(* IEC 61131-3 sources: kns-pump-station/tests/POUs/Station/FB_Protections_Test, 24 files *)

(* ---- DryRunAndEmergencyBothDryRunWins.method.decl.st ---- *)
// 04 §10.2: сухой ход и аварийный уровень одновременно — оба признака (старшинство сухого хода —
// FB_ControlSelector), по поплавкам LS103 останавливает откачку
METHOD PRIVATE DryRunAndEmergencyBothDryRunWins
VAR
    fbDut  : FB_Protections;            // ФБ под тестом
    fbTime : PL.FB_FakeTime;            // подменное время, старт 1 ч
    stCfg  : ST_StationCfg;             // уставки по умолчанию (tLdev 30 с, tLtRecover 30 с, tDryRelease 60 с)
    fbSink : FB_FakeEventSink;          // подменный журнал
END_VAR

(* ---- DryRunByFloat.method.decl.st ---- *)
// 04 §10.1, PMI-19: поплавок LS103 сработал — сухой ход сразу (защита срабатывает до проверки согласования)
METHOD PRIVATE DryRunByFloat
VAR
    fbDut  : FB_Protections;            // ФБ под тестом
    fbTime : PL.FB_FakeTime;            // подменное время, старт 1 ч
    stCfg  : ST_StationCfg;             // уставки по умолчанию (tLdev 30 с, tLtRecover 30 с, tDryRelease 60 с)
    fbSink : FB_FakeEventSink;          // подменный журнал
END_VAR

(* ---- DryRunByLtLl.method.decl.st ---- *)
// 04 §10.1, PMI-18: LL по годному уровнемеру — сухой ход
METHOD PRIVATE DryRunByLtLl
VAR
    fbDut  : FB_Protections;            // ФБ под тестом
    fbTime : PL.FB_FakeTime;            // подменное время, старт 1 ч
    stCfg  : ST_StationCfg;             // уставки по умолчанию (tLdev 30 с, tLtRecover 30 с, tDryRelease 60 с)
    fbSink : FB_FakeEventSink;          // подменный журнал
END_VAR

(* ---- DryRunReleaseAboveL.method.decl.st ---- *)
// 04 §10.1, PMI-18: снятие сухого хода — LS103 не сработал, нет LL и уровень выше L (по флагу L уровнемера)
METHOD PRIVATE DryRunReleaseAboveL
VAR
    fbDut  : FB_Protections;            // ФБ под тестом
    fbTime : PL.FB_FakeTime;            // подменное время, старт 1 ч
    stCfg  : ST_StationCfg;             // уставки по умолчанию (tLdev 30 с, tLtRecover 30 с, tDryRelease 60 с)
    fbSink : FB_FakeEventSink;          // подменный журнал
END_VAR

(* ---- DryRunReleaseWithoutLtAfterTDryRelease.method.decl.st ---- *)
// 04 §10.1, §11, PMI-19: без уровнемера сухой ход снимается, когда LS103 снят дольше tDryRelease = 60 с (не
// раньше)
METHOD PRIVATE DryRunReleaseWithoutLtAfterTDryRelease
VAR
    fbDut  : FB_Protections;            // ФБ под тестом
    fbTime : PL.FB_FakeTime;            // подменное время, старт 1 ч
    stCfg  : ST_StationCfg;             // уставки по умолчанию (tLdev 30 с, tLtRecover 30 с, tDryRelease 60 с)
    fbSink : FB_FakeEventSink;          // подменный журнал
END_VAR

(* ---- EmergencyByFloatAndByHh.method.decl.st ---- *)
// 04 §10.2, PMI-20, PMI-23: аварийный уровень — по LS102 и по HH годного уровнемера
METHOD PRIVATE EmergencyByFloatAndByHh
VAR
    fbDut  : FB_Protections;            // ФБ под тестом
    fbTime : PL.FB_FakeTime;            // подменное время, старт 1 ч
    stCfg  : ST_StationCfg;             // уставки по умолчанию (tLdev 30 с, tLtRecover 30 с, tDryRelease 60 с)
    fbSink : FB_FakeEventSink;          // подменный журнал
    fbDut2 : FB_Protections;           // второй экземпляр: HH
END_VAR

(* ---- EmergencyReleaseBelowH.method.decl.st ---- *)
// 04 §10.2, PMI-20: снятие аварийного режима — LS102 снят и уровень ниже H
METHOD PRIVATE EmergencyReleaseBelowH
VAR
    fbDut  : FB_Protections;            // ФБ под тестом
    fbTime : PL.FB_FakeTime;            // подменное время, старт 1 ч
    stCfg  : ST_StationCfg;             // уставки по умолчанию (tLdev 30 с, tLtRecover 30 с, tDryRelease 60 с)
    fbSink : FB_FakeEventSink;          // подменный журнал
END_VAR

(* ---- FalseLs102MaskedAfterTLdev.method.decl.st ---- *)
// 04 §10.5, PMI-23: LS102 сработал при уровне ниже 3,50 м — через tLdev поплавок исключён (101011, 102), аварийный
// режим снят
METHOD PRIVATE FalseLs102MaskedAfterTLdev
VAR
    fbDut  : FB_Protections;            // ФБ под тестом
    fbTime : PL.FB_FakeTime;            // подменное время, старт 1 ч
    stCfg  : ST_StationCfg;             // уставки по умолчанию (tLdev 30 с, tLtRecover 30 с, tDryRelease 60 с)
    fbSink : FB_FakeEventSink;          // подменный журнал
END_VAR

(* ---- FalseLs103MaskedAfterTLdev.method.decl.st ---- *)
// 04 §10.5, PMI-22: LS103 сработал при уровне выше 0,80 м и уровнемере в норме — через tLdev поплавок исключён
// (101011, 103), KNS1.LDEV, сухой ход снят
METHOD PRIVATE FalseLs103MaskedAfterTLdev
VAR
    fbDut  : FB_Protections;            // ФБ под тестом
    fbTime : PL.FB_FakeTime;            // подменное время, старт 1 ч
    stCfg  : ST_StationCfg;             // уставки по умолчанию (tLdev 30 с, tLtRecover 30 с, tDryRelease 60 с)
    fbSink : FB_FakeEventSink;          // подменный журнал
END_VAR

(* ---- FirstCallDoesNotEnterFloatMode.method.decl.st ---- *)
// DESIGN 7: в первом цикле выходы устройств ещё не посчитаны (xValid = FALSE) — режим по поплавкам не включается
METHOD PRIVATE FirstCallDoesNotEnterFloatMode
VAR
    fbDut  : FB_Protections;            // ФБ под тестом
    fbTime : PL.FB_FakeTime;            // подменное время, старт 1 ч
    stCfg  : ST_StationCfg;             // уставки по умолчанию (tLdev 30 с, tLtRecover 30 с, tDryRelease 60 с)
    fbSink : FB_FakeEventSink;          // подменный журнал
END_VAR

(* ---- FloatModeEntryWhilePumpingKeepsPumping.method.decl.st ---- *)
// 04 §11, PMI-25: отказ уровнемера при работающих насосах — сразу «откачка» до LS103
METHOD PRIVATE FloatModeEntryWhilePumpingKeepsPumping
VAR
    fbDut  : FB_Protections;            // ФБ под тестом
    fbTime : PL.FB_FakeTime;            // подменное время, старт 1 ч
    stCfg  : ST_StationCfg;             // уставки по умолчанию (tLdev 30 с, tLtRecover 30 с, tDryRelease 60 с)
    fbSink : FB_FakeEventSink;          // подменный журнал
END_VAR

(* ---- FloatModeExitAfterTLtRecover.method.decl.st ---- *)
// 04 §11, PMI-27: уровнемер снова годен — режим по поплавкам ещё tLtRecover = 30 с, затем выход (101014)
METHOD PRIVATE FloatModeExitAfterTLtRecover
VAR
    fbDut  : FB_Protections;            // ФБ под тестом
    fbTime : PL.FB_FakeTime;            // подменное время, старт 1 ч
    stCfg  : ST_StationCfg;             // уставки по умолчанию (tLdev 30 с, tLtRecover 30 с, tDryRelease 60 с)
    fbSink : FB_FakeEventSink;          // подменный журнал
END_VAR

(* ---- FloatModeStartsAllOnLs102StopsOnLs103.method.decl.st ---- *)
// 04 §11, PMI-21, PMI-25: по поплавкам — ожидание LS102, затем откачка всеми насосами до LS103
METHOD PRIVATE FloatModeStartsAllOnLs102StopsOnLs103
VAR
    fbDut  : FB_Protections;            // ФБ под тестом
    fbTime : PL.FB_FakeTime;            // подменное время, старт 1 ч
    stCfg  : ST_StationCfg;             // уставки по умолчанию (tLdev 30 с, tLtRecover 30 с, tDryRelease 60 с)
    fbSink : FB_FakeEventSink;          // подменный журнал
END_VAR

(* ---- GoodLtContradictingFloatMasksFloat.method.decl.st ---- *)
// 04 §10.5: при уровнемере в норме (Good) виноват поплавок — исключается поплавок, уровнемер остаётся в логике
METHOD PRIVATE GoodLtContradictingFloatMasksFloat
VAR
    fbDut  : FB_Protections;            // ФБ под тестом
    fbTime : PL.FB_FakeTime;            // подменное время, старт 1 ч
    stCfg  : ST_StationCfg;             // уставки по умолчанию (tLdev 30 с, tLtRecover 30 с, tDryRelease 60 с)
    fbSink : FB_FakeEventSink;          // подменный журнал
END_VAR

(* ---- Ls102NotTrippedAboveOffMark.method.decl.st ---- *)
// 04 §10.5, PMI-24: LS102 не сработал при уровне выше 4,40 м — через tLdev KNS1.LDEV; аварийный режим держит HH
// уровнемера, маски нет
METHOD PRIVATE Ls102NotTrippedAboveOffMark
VAR
    fbDut  : FB_Protections;            // ФБ под тестом
    fbTime : PL.FB_FakeTime;            // подменное время, старт 1 ч
    stCfg  : ST_StationCfg;             // уставки по умолчанию (tLdev 30 с, tLtRecover 30 с, tDryRelease 60 с)
    fbSink : FB_FakeEventSink;          // подменный журнал
END_VAR

(* ---- Ls103NotTrippedBelowOffMark.method.decl.st ---- *)
// 04 §10.5: LS103 не сработал при уровне ниже 0,20 м и уровнемере в норме — через tLdev KNS1.LDEV, защиту держит
// LL уровнемера
METHOD PRIVATE Ls103NotTrippedBelowOffMark
VAR
    fbDut  : FB_Protections;            // ФБ под тестом
    fbTime : PL.FB_FakeTime;            // подменное время, старт 1 ч
    stCfg  : ST_StationCfg;             // уставки по умолчанию (tLdev 30 с, tLtRecover 30 с, tDryRelease 60 с)
    fbSink : FB_FakeEventSink;          // подменный журнал
END_VAR

(* ---- MaskReleasedWhenFloatReturns.method.decl.st ---- *)
// 04 §10.5, PMI-22 шаг 2: маска снимается сама, когда поплавок вернулся (101012, 103)
METHOD PRIVATE MaskReleasedWhenFloatReturns
VAR
    fbDut  : FB_Protections;            // ФБ под тестом
    fbTime : PL.FB_FakeTime;            // подменное время, старт 1 ч
    stCfg  : ST_StationCfg;             // уставки по умолчанию (tLdev 30 с, tLtRecover 30 с, tDryRelease 60 с)
    fbSink : FB_FakeEventSink;          // подменный журнал
END_VAR

(* ---- MaskReleasedWhenLtInvalid.method.decl.st ---- *)
// 04 §10.5: маска поплавка снимается сразу, когда уровнемер стал негоден: поплавок снова защищает (сухой ход)
METHOD PRIVATE MaskReleasedWhenLtInvalid
VAR
    fbDut  : FB_Protections;            // ФБ под тестом
    fbTime : PL.FB_FakeTime;            // подменное время, старт 1 ч
    stCfg  : ST_StationCfg;             // уставки по умолчанию (tLdev 30 с, tLtRecover 30 с, tDryRelease 60 с)
    fbSink : FB_FakeEventSink;          // подменный журнал
END_VAR

(* ---- OorLtInvalidFloatsAtOnce.method.decl.st ---- *)
// 04 §10.5, §11, PMI-26, AI-13 plc-process-lib 1.0.0: настоящий PL.FB_AnalogInput с уставками LT101 проекта.
// Ток 3,7 мА (выход за диапазон без отказа): до подтверждения (tFailDelay 2 с) значение годно, сухого хода нет;
// после — xValid = FALSE и NE 107 «вне спецификации»: сразу режим по поплавкам (101013). Уставки считаются по
// значению насыщения (LL уровнемера есть), но сухого хода по уровнемеру нет, противоречие с LS103 не считается
// (KNS1.LDEV нет): защиту держит поплавок
METHOD PRIVATE OorLtInvalidFloatsAtOnce
VAR
    fbDut   : FB_Protections;           // ФБ под тестом
    fbTime  : PL.FB_FakeTime;           // подменное время, старт 1 ч
    stCfg   : ST_StationCfg;            // уставки по умолчанию (tLdev 30 с)
    fbSink  : FB_FakeEventSink;         // подменный журнал
    stAiCmd : PL.ST_AnalogInputCmd;     // GVL_Hmi.stLT101Cmd
    stAiCfg : PL.ST_AnalogInputCfg;     // GVL_Persist.stLT101Cfg — уставки проекта
END_VAR
VAR_INST
    fbLT101 : PL.FB_AnalogInput;        // GVL_Devices.fbLT101
END_VAR

(* ---- Run.method.decl.st ---- *)
// Помощник: uiSteps шагов времени tStep; входы ФБ тест задаёт присваиванием до вызова
METHOD PRIVATE Run
VAR_IN_OUT
    fbDut  : FB_Protections;            // ФБ под тестом
    fbTime : PL.FB_FakeTime;            // подменное время
    stCfg  : ST_StationCfg;             // уставки
END_VAR
VAR_INPUT
    tStep   : TIME;                     // шаг времени
    uiSteps : UINT;                     // шагов
END_VAR
VAR
    uiStep : UINT;                      // номер шага
END_VAR

(* ---- Run.method.impl.st ---- *)
FOR uiStep := 1 TO uiSteps DO
    fbTime.Advance(tStep := tStep);
    fbDut(itfTime := fbTime, stCfg := stCfg);
END_FOR

(* ---- RunWithAi.method.decl.st ---- *)
// Помощник: uiSteps шагов по 100 мс — настоящий уровнемер PL.FB_AnalogInput (ток rIn_mA), затем FB_Protections
// с его выходами, как в PRG_Station (уровень, xValid, NE 107, уставки L, LL, H, HH)
METHOD PRIVATE RunWithAi
VAR_IN_OUT
    fbDut   : FB_Protections;           // ФБ под тестом
    fbTime  : PL.FB_FakeTime;           // подменное время
    stCfg   : ST_StationCfg;            // уставки станции
    fbAi    : PL.FB_AnalogInput;        // GVL_Devices.fbLT101
    stAiCmd : PL.ST_AnalogInputCmd;     // GVL_Hmi.stLT101Cmd
    stAiCfg : PL.ST_AnalogInputCfg;     // GVL_Persist.stLT101Cfg
END_VAR
VAR_INPUT
    rIn_mA  : REAL;                     // ток LT101
    uiSteps : UINT;                     // шагов по 100 мс
END_VAR
VAR
    uiStep : UINT;                      // номер шага
END_VAR

(* ---- RunWithAi.method.impl.st ---- *)
FOR uiStep := 1 TO uiSteps DO
    fbTime.Advance(tStep := T#100MS);
    fbAi(rIn := rIn_mA, xChannelFault := FALSE, itfTime := fbTime, stCmd := stAiCmd, stCfg := stAiCfg);
    fbDut.rLevel_m := fbAi.rValue_eu;
    fbDut.xLevelValid := fbAi.xValid;
    fbDut.eLevelNe107 := fbAi.stSts.stCommon.eNe107;
    fbDut.xLevelL := fbAi.xL;
    fbDut.xLevelLL := fbAi.xLL;
    fbDut.xLevelH := fbAi.xH;
    fbDut.xLevelHH := fbAi.xHH;
    fbDut(itfTime := fbTime, stCfg := stCfg);
END_FOR

(* ---- TimeBackwardsRestartsLdev.method.decl.st ---- *)
// Время назад — выдержка tLdev контроля согласования начинается заново, поплавок раньше срока не исключается
METHOD PRIVATE TimeBackwardsRestartsLdev
VAR
    fbDut  : FB_Protections;            // ФБ под тестом
    fbTime : PL.FB_FakeTime;            // подменное время, старт 1 ч
    stCfg  : ST_StationCfg;             // уставки по умолчанию (tLdev 30 с, tLtRecover 30 с, tDryRelease 60 с)
    fbSink : FB_FakeEventSink;          // подменный журнал
END_VAR
